// TIA Portal V17 export
// export: Created 2025-07-10T12:23:13.1481267Z, ExportSetting WithDefaults, DisplayName Totally Integrated Automation Portal, DisplayVersion V17, DisplayName TIA Portal Openness, DisplayVersion V17, DisplayName TIA Portal Version Control Interface, DisplayVersion V17, DisplayName SINAMICS Startdrive Advanced, DisplayVersion V17, DisplayName SINAMICS Startdrive G130, G150, S120, S150, SINAMICS MV, S210, DisplayVersion V17, DisplayName SINAMICS Startdrive G110M, G120, G120C, G120D, G120P, G115D, DisplayVersion V17, DisplayName STEP 7 Professional, DisplayVersion V17, DisplayName STEP 7 Safety, DisplayVersion V17, DisplayName WinCC Professional, DisplayVersion V17
FUNCTION_BLOCK "PR_PC4005_Operator_DecisionV4_77a371"   // FB1, LAD
VERSION : 0.1
// stored: AutoNumber true, IsIECCheckEnabled false, UDAEnableTagReadback false
   VAR_INPUT
      iAutoRunning : Bool;
      iOperatorAuthorizationPB : Bool;
      iPCAckZero : Bool;
      iPCBypass : Bool;
      iPCDataReadOver : Bool;
      iPCDataWriteOver : Bool;
      iPalletPresentAtStation : Bool;
      iProcessOver : Bool;
      iProcessStartFormPZR : Bool;
      iRejectPB : Bool;
      iResetMem : Bool;
      iReset_fault : Bool;
      iScanOver : Bool;
      iScanResultNok : Bool;
      iScanResultOk : Bool;
      iScannerBypass : Bool;
      iSstMode : Bool;
      iSstPB : Bool;
      iUnloadCycleSelection : Bool;
   END_VAR
   VAR_OUTPUT
      qPCReadCmd : Bool;
      qPCWriteCmd : Bool;
      qProcessOver : Bool;
      qResetPalletStatusData : Bool;
      qScanCmd : Bool;
   END_VAR
   VAR DB_SPECIFIC
      StateNo : Int;
      s29_WaitProcStart : Bool;
      s29_WaitProcStart_T1 : Bool;
      s30_WaitCartnSheetOp : Bool;
      s30_WaitCartnSheetOp_T1 : Bool;
      s31_ChkCycleSelect : Bool;
      s31_ChkCycleSelect_T1 : Bool;
      s31_ChkCycleSelect_T2 : Bool;
      s32_WaitScanOver : Bool;
      s32_WaitScanOver_T1 : Bool;
      s33_ChkScanResult : Bool;
      s33_ChkScanResult_T1 : Bool;
      s33_ChkScanResult_T2 : Bool;
      s34_WaitOpDecision : Bool;
      s34_WaitOpDecision_T1 : Bool;
      s34_WaitOpDecision_T2 : Bool;
      s35_ChkPCAckReset0 : Bool;
      s35_ChkPCAckReset0_T1 : Bool;
      s36_WaitDataReadPC : Bool;
      s36_WaitDataReadPC_T1 : Bool;
      s38_WaitProcStartLow : Bool;
      s38_WaitProcStartLow_T1 : Bool;
      s39_WaitPalletAbsnt : Bool;
      s39_WaitPalletAbsnt_T1 : Bool;
      s40_WaitFaultReset : Bool;
      s40_WaitFaultReset_T1 : Bool;
      s41_ChkPCAckReset0Up : Bool;
      s41_ChkPCAckReset0Up_T1 : Bool;
      s42_WaitDataUploadPC : Bool;
      s42_WaitDataUploadPC_T1 : Bool;
      s43_ChkRecovery : Bool;
      s43_ChkRecovery_T1 : Bool;
      s43_ChkRecovery_T2 : Bool;
      sPalletAccepted : Bool;
      sProcessOver : Bool;
      sSst : Bool;
      sSstPulse : Bool;
      sSstRise : Bool;
      sStWtResetRel : Bool;
      sStWtResetRel_T1 : Bool;
   END_VAR
   VAR_TEMP
      tOne : Bool;
   END_VAR
   VAR_TEMP   // added for the SCL form of the ladder/FBD networks
      _w1 : Bool;
   END_VAR
BEGIN

REGION Network 1
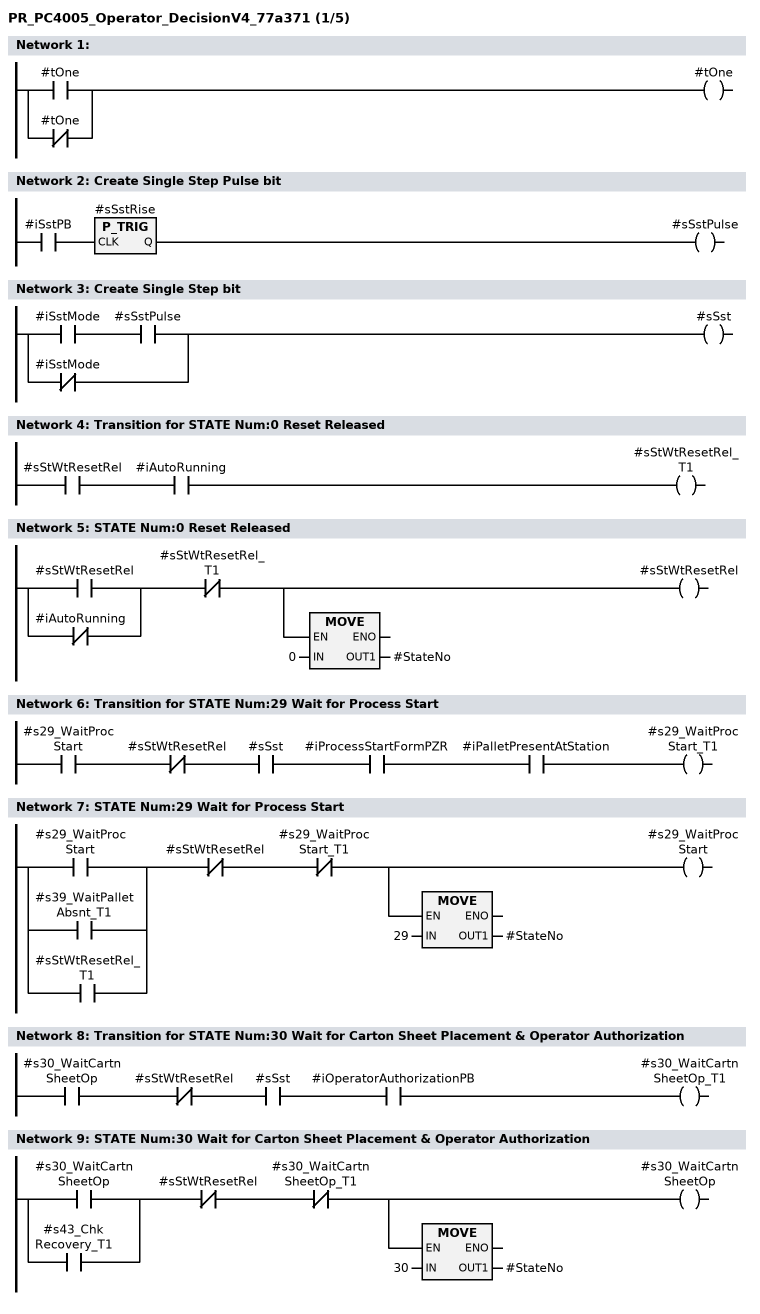
   RUNG wire#powerrail
      Contact( #tOne )
      wire#w1
      Coil( #tOne )
   END_RUNG
   RUNG wire#powerrail
      I_Contact( #tOne )
   END_RUNG wire#w1
   // the same network as SCL:
   #tOne := #tOne OR NOT #tOne;
END_REGION

REGION Network 2: Create Single Step Pulse bit
   RUNG wire#powerrail
      Contact( #iSstPB )
      P_Trig( #sSstRise )
      Coil( #sSstPulse )
   END_RUNG
   // the same network as SCL:
   #_w1 := #iSstPB AND NOT #sSstRise;   // rising edge
   #sSstRise := #iSstPB;
   #sSstPulse := #_w1;
END_REGION

REGION Network 3: Create Single Step bit
   RUNG wire#powerrail
      Contact( #iSstMode )
      Contact( #sSstPulse )
      wire#w1
      Coil( #sSst )
   END_RUNG
   RUNG wire#powerrail
      I_Contact( #iSstMode )
   END_RUNG wire#w1
   // the same network as SCL:
   #sSst := (#iSstMode AND #sSstPulse) OR NOT #iSstMode;
END_REGION

REGION Network 4: Transition for STATE Num:0 Reset Released
   RUNG wire#powerrail
      Contact( #sStWtResetRel )
      Contact( #iAutoRunning )
      Coil( #sStWtResetRel_T1 )
   END_RUNG
   // the same network as SCL:
   #sStWtResetRel_T1 := #sStWtResetRel AND #iAutoRunning;
END_REGION

REGION Network 5: STATE Num:0 Reset Released
   RUNG wire#powerrail
      Contact( #sStWtResetRel )
      wire#w1
      I_Contact( #sStWtResetRel_T1 )
      wire#w2
      Coil( #sStWtResetRel )
   END_RUNG
   RUNG wire#powerrail
      I_Contact( #iAutoRunning )
   END_RUNG wire#w1
   RUNG wire#w2
      { S7_GenerateENO := "TRUE" } Move(in := 0, out1 => #StateNo)
   END_RUNG
   // the same network as SCL:
   #sStWtResetRel := (#sStWtResetRel OR NOT #iAutoRunning) AND NOT #sStWtResetRel_T1;
   IF #sStWtResetRel THEN #StateNo := 0; END_IF;
END_REGION

REGION Network 6: Transition for STATE Num:29 Wait for Process Start
   RUNG wire#powerrail
      Contact( #s29_WaitProcStart )
      I_Contact( #sStWtResetRel )
      Contact( #sSst )
      Contact( #iProcessStartFormPZR )
      Contact( #iPalletPresentAtStation )
      Coil( #s29_WaitProcStart_T1 )
   END_RUNG
   // the same network as SCL:
   #s29_WaitProcStart_T1 := #s29_WaitProcStart AND NOT #sStWtResetRel AND #sSst AND #iProcessStartFormPZR AND #iPalletPresentAtStation;
END_REGION

REGION Network 7: STATE Num:29 Wait for Process Start
   RUNG wire#powerrail
      Contact( #s29_WaitProcStart )
      wire#w1
      I_Contact( #sStWtResetRel )
      I_Contact( #s29_WaitProcStart_T1 )
      wire#w2
      Coil( #s29_WaitProcStart )
   END_RUNG
   RUNG wire#powerrail
      Contact( #s39_WaitPalletAbsnt_T1 )
   END_RUNG wire#w1
   RUNG wire#powerrail
      Contact( #sStWtResetRel_T1 )
   END_RUNG wire#w1
   RUNG wire#w2
      { S7_GenerateENO := "TRUE" } Move(in := 29, out1 => #StateNo)
   END_RUNG
   // the same network as SCL:
   #s29_WaitProcStart := (#s29_WaitProcStart OR #s39_WaitPalletAbsnt_T1 OR #sStWtResetRel_T1) AND NOT #sStWtResetRel AND NOT #s29_WaitProcStart_T1;
   IF #s29_WaitProcStart THEN #StateNo := 29; END_IF;
END_REGION

REGION Network 8: Transition for STATE Num:30 Wait for Carton Sheet Placement & Operator Authorization
   RUNG wire#powerrail
      Contact( #s30_WaitCartnSheetOp )
      I_Contact( #sStWtResetRel )
      Contact( #sSst )
      Contact( #iOperatorAuthorizationPB )
      Coil( #s30_WaitCartnSheetOp_T1 )
   END_RUNG
   // the same network as SCL:
   #s30_WaitCartnSheetOp_T1 := #s30_WaitCartnSheetOp AND NOT #sStWtResetRel AND #sSst AND #iOperatorAuthorizationPB;
END_REGION

REGION Network 9: STATE Num:30 Wait for Carton Sheet Placement & Operator Authorization
   RUNG wire#powerrail
      Contact( #s30_WaitCartnSheetOp )
      wire#w1
      I_Contact( #sStWtResetRel )
      I_Contact( #s30_WaitCartnSheetOp_T1 )
      wire#w2
      Coil( #s30_WaitCartnSheetOp )
   END_RUNG
   RUNG wire#powerrail
      Contact( #s43_ChkRecovery_T1 )
   END_RUNG wire#w1
   RUNG wire#w2
      { S7_GenerateENO := "TRUE" } Move(in := 30, out1 => #StateNo)
   END_RUNG
   // the same network as SCL:
   #s30_WaitCartnSheetOp := (#s30_WaitCartnSheetOp OR #s43_ChkRecovery_T1) AND NOT #sStWtResetRel AND NOT #s30_WaitCartnSheetOp_T1;
   IF #s30_WaitCartnSheetOp THEN #StateNo := 30; END_IF;
END_REGION

REGION Network 10: Transition for STATE Num:31 Check Cycle Selection
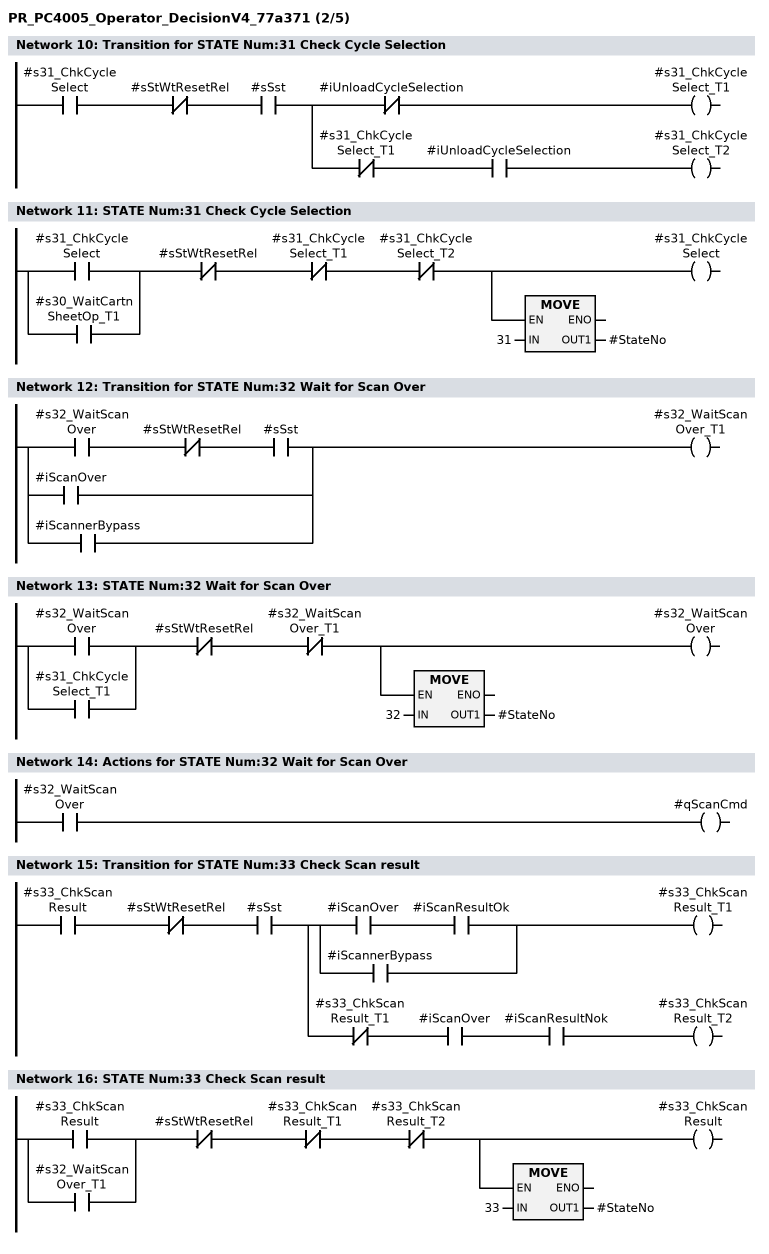
   RUNG wire#powerrail
      Contact( #s31_ChkCycleSelect )
      I_Contact( #sStWtResetRel )
      Contact( #sSst )
      wire#w1
      I_Contact( #iUnloadCycleSelection )
      Coil( #s31_ChkCycleSelect_T1 )
   END_RUNG
   RUNG wire#w1
      I_Contact( #s31_ChkCycleSelect_T1 )
      Contact( #iUnloadCycleSelection )
      Coil( #s31_ChkCycleSelect_T2 )
   END_RUNG
   // the same network as SCL:
   #_w1 := #s31_ChkCycleSelect AND NOT #sStWtResetRel AND #sSst;
   #s31_ChkCycleSelect_T1 := #_w1 AND NOT #iUnloadCycleSelection;
   #s31_ChkCycleSelect_T2 := #_w1 AND NOT #s31_ChkCycleSelect_T1 AND #iUnloadCycleSelection;
END_REGION

REGION Network 11: STATE Num:31 Check Cycle Selection
   RUNG wire#powerrail
      Contact( #s31_ChkCycleSelect )
      wire#w1
      I_Contact( #sStWtResetRel )
      I_Contact( #s31_ChkCycleSelect_T1 )
      I_Contact( #s31_ChkCycleSelect_T2 )
      wire#w2
      Coil( #s31_ChkCycleSelect )
   END_RUNG
   RUNG wire#powerrail
      Contact( #s30_WaitCartnSheetOp_T1 )
   END_RUNG wire#w1
   RUNG wire#w2
      { S7_GenerateENO := "TRUE" } Move(in := 31, out1 => #StateNo)
   END_RUNG
   // the same network as SCL:
   #s31_ChkCycleSelect := (#s31_ChkCycleSelect OR #s30_WaitCartnSheetOp_T1) AND NOT #sStWtResetRel AND NOT #s31_ChkCycleSelect_T1 AND NOT #s31_ChkCycleSelect_T2;
   IF #s31_ChkCycleSelect THEN #StateNo := 31; END_IF;
END_REGION

REGION Network 12: Transition for STATE Num:32 Wait for Scan Over
   RUNG wire#powerrail
      Contact( #s32_WaitScanOver )
      I_Contact( #sStWtResetRel )
      Contact( #sSst )
      wire#w1
      Coil( #s32_WaitScanOver_T1 )
   END_RUNG
   RUNG wire#powerrail
      Contact( #iScanOver )
   END_RUNG wire#w1
   RUNG wire#powerrail
      Contact( #iScannerBypass )
   END_RUNG wire#w1
   // the same network as SCL:
   #s32_WaitScanOver_T1 := (#s32_WaitScanOver AND NOT #sStWtResetRel AND #sSst) OR #iScanOver OR #iScannerBypass;
END_REGION

REGION Network 13: STATE Num:32 Wait for Scan Over
   RUNG wire#powerrail
      Contact( #s32_WaitScanOver )
      wire#w1
      I_Contact( #sStWtResetRel )
      I_Contact( #s32_WaitScanOver_T1 )
      wire#w2
      Coil( #s32_WaitScanOver )
   END_RUNG
   RUNG wire#powerrail
      Contact( #s31_ChkCycleSelect_T1 )
   END_RUNG wire#w1
   RUNG wire#w2
      { S7_GenerateENO := "TRUE" } Move(in := 32, out1 => #StateNo)
   END_RUNG
   // the same network as SCL:
   #s32_WaitScanOver := (#s32_WaitScanOver OR #s31_ChkCycleSelect_T1) AND NOT #sStWtResetRel AND NOT #s32_WaitScanOver_T1;
   IF #s32_WaitScanOver THEN #StateNo := 32; END_IF;
END_REGION

REGION Network 14: Actions for STATE Num:32 Wait for Scan Over
   RUNG wire#powerrail
      Contact( #s32_WaitScanOver )
      Coil( #qScanCmd )
   END_RUNG
   // the same network as SCL:
   #qScanCmd := #s32_WaitScanOver;
END_REGION

REGION Network 15: Transition for STATE Num:33 Check Scan result
   RUNG wire#powerrail
      Contact( #s33_ChkScanResult )
      I_Contact( #sStWtResetRel )
      Contact( #sSst )
      wire#w1
      Contact( #iScanOver )
      Contact( #iScanResultOk )
      wire#w2
      Coil( #s33_ChkScanResult_T1 )
   END_RUNG
   RUNG wire#w1
      Contact( #iScannerBypass )
   END_RUNG wire#w2
   RUNG wire#w1
      I_Contact( #s33_ChkScanResult_T1 )
      Contact( #iScanOver )
      Contact( #iScanResultNok )
      Coil( #s33_ChkScanResult_T2 )
   END_RUNG
   // the same network as SCL:
   #_w1 := #s33_ChkScanResult AND NOT #sStWtResetRel AND #sSst;
   #s33_ChkScanResult_T1 := #_w1 AND ((#iScanOver AND #iScanResultOk) OR #iScannerBypass);
   #s33_ChkScanResult_T2 := #_w1 AND NOT #s33_ChkScanResult_T1 AND #iScanOver AND #iScanResultNok;
END_REGION

REGION Network 16: STATE Num:33 Check Scan result
   RUNG wire#powerrail
      Contact( #s33_ChkScanResult )
      wire#w1
      I_Contact( #sStWtResetRel )
      I_Contact( #s33_ChkScanResult_T1 )
      I_Contact( #s33_ChkScanResult_T2 )
      wire#w2
      Coil( #s33_ChkScanResult )
   END_RUNG
   RUNG wire#powerrail
      Contact( #s32_WaitScanOver_T1 )
   END_RUNG wire#w1
   RUNG wire#w2
      { S7_GenerateENO := "TRUE" } Move(in := 33, out1 => #StateNo)
   END_RUNG
   // the same network as SCL:
   #s33_ChkScanResult := (#s33_ChkScanResult OR #s32_WaitScanOver_T1) AND NOT #sStWtResetRel AND NOT #s33_ChkScanResult_T1 AND NOT #s33_ChkScanResult_T2;
   IF #s33_ChkScanResult THEN #StateNo := 33; END_IF;
END_REGION

REGION Network 17: Transition for STATE Num:34 Wait for Operator Decision
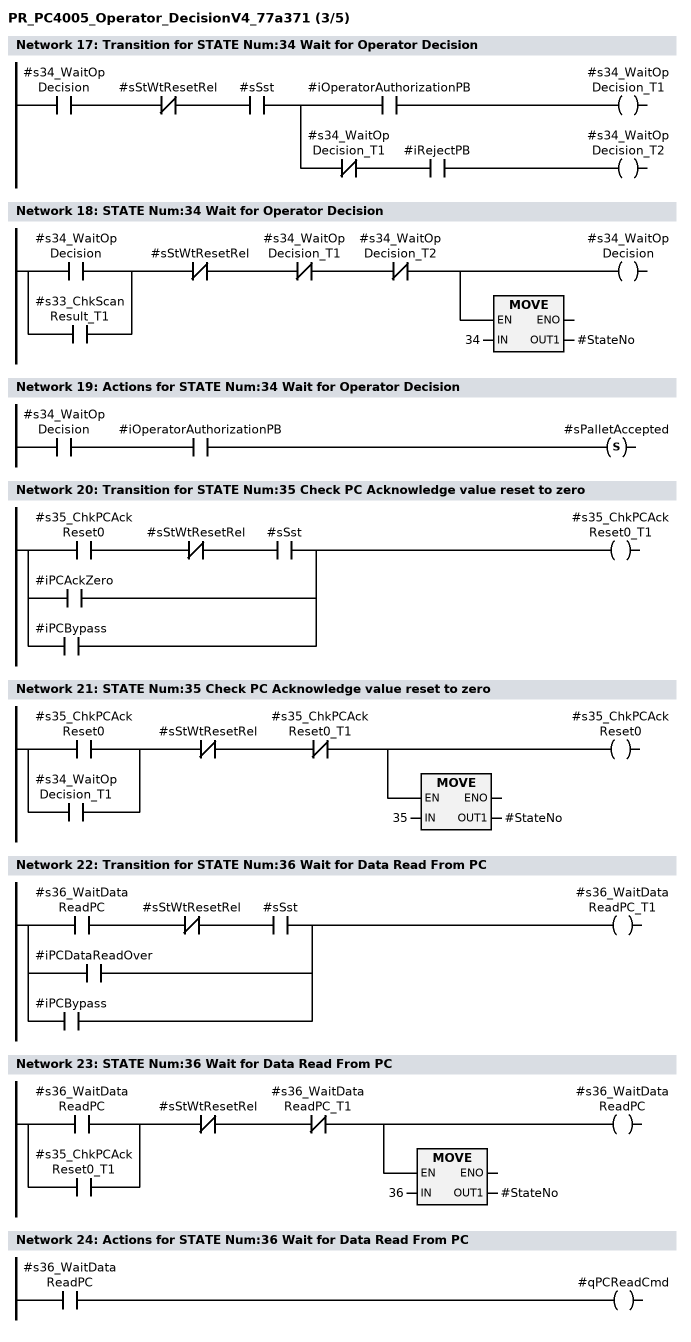
   RUNG wire#powerrail
      Contact( #s34_WaitOpDecision )
      I_Contact( #sStWtResetRel )
      Contact( #sSst )
      wire#w1
      Contact( #iOperatorAuthorizationPB )
      Coil( #s34_WaitOpDecision_T1 )
   END_RUNG
   RUNG wire#w1
      I_Contact( #s34_WaitOpDecision_T1 )
      Contact( #iRejectPB )
      Coil( #s34_WaitOpDecision_T2 )
   END_RUNG
   // the same network as SCL:
   #_w1 := #s34_WaitOpDecision AND NOT #sStWtResetRel AND #sSst;
   #s34_WaitOpDecision_T1 := #_w1 AND #iOperatorAuthorizationPB;
   #s34_WaitOpDecision_T2 := #_w1 AND NOT #s34_WaitOpDecision_T1 AND #iRejectPB;
END_REGION

REGION Network 18: STATE Num:34 Wait for Operator Decision
   RUNG wire#powerrail
      Contact( #s34_WaitOpDecision )
      wire#w1
      I_Contact( #sStWtResetRel )
      I_Contact( #s34_WaitOpDecision_T1 )
      I_Contact( #s34_WaitOpDecision_T2 )
      wire#w2
      Coil( #s34_WaitOpDecision )
   END_RUNG
   RUNG wire#powerrail
      Contact( #s33_ChkScanResult_T1 )
   END_RUNG wire#w1
   RUNG wire#w2
      { S7_GenerateENO := "TRUE" } Move(in := 34, out1 => #StateNo)
   END_RUNG
   // the same network as SCL:
   #s34_WaitOpDecision := (#s34_WaitOpDecision OR #s33_ChkScanResult_T1) AND NOT #sStWtResetRel AND NOT #s34_WaitOpDecision_T1 AND NOT #s34_WaitOpDecision_T2;
   IF #s34_WaitOpDecision THEN #StateNo := 34; END_IF;
END_REGION

REGION Network 19: Actions for STATE Num:34 Wait for Operator Decision
   RUNG wire#powerrail
      Contact( #s34_WaitOpDecision )
      Contact( #iOperatorAuthorizationPB )
      S_Coil( #sPalletAccepted )
   END_RUNG
   // the same network as SCL:
   IF #s34_WaitOpDecision AND #iOperatorAuthorizationPB THEN #sPalletAccepted := TRUE; END_IF;
END_REGION

REGION Network 20: Transition for STATE Num:35 Check PC Acknowledge value reset to zero
   RUNG wire#powerrail
      Contact( #s35_ChkPCAckReset0 )
      I_Contact( #sStWtResetRel )
      Contact( #sSst )
      wire#w1
      Coil( #s35_ChkPCAckReset0_T1 )
   END_RUNG
   RUNG wire#powerrail
      Contact( #iPCAckZero )
   END_RUNG wire#w1
   RUNG wire#powerrail
      Contact( #iPCBypass )
   END_RUNG wire#w1
   // the same network as SCL:
   #s35_ChkPCAckReset0_T1 := (#s35_ChkPCAckReset0 AND NOT #sStWtResetRel AND #sSst) OR #iPCAckZero OR #iPCBypass;
END_REGION

REGION Network 21: STATE Num:35 Check PC Acknowledge value reset to zero
   RUNG wire#powerrail
      Contact( #s35_ChkPCAckReset0 )
      wire#w1
      I_Contact( #sStWtResetRel )
      I_Contact( #s35_ChkPCAckReset0_T1 )
      wire#w2
      Coil( #s35_ChkPCAckReset0 )
   END_RUNG
   RUNG wire#powerrail
      Contact( #s34_WaitOpDecision_T1 )
   END_RUNG wire#w1
   RUNG wire#w2
      { S7_GenerateENO := "TRUE" } Move(in := 35, out1 => #StateNo)
   END_RUNG
   // the same network as SCL:
   #s35_ChkPCAckReset0 := (#s35_ChkPCAckReset0 OR #s34_WaitOpDecision_T1) AND NOT #sStWtResetRel AND NOT #s35_ChkPCAckReset0_T1;
   IF #s35_ChkPCAckReset0 THEN #StateNo := 35; END_IF;
END_REGION

REGION Network 22: Transition for STATE Num:36 Wait for Data Read From PC
   RUNG wire#powerrail
      Contact( #s36_WaitDataReadPC )
      I_Contact( #sStWtResetRel )
      Contact( #sSst )
      wire#w1
      Coil( #s36_WaitDataReadPC_T1 )
   END_RUNG
   RUNG wire#powerrail
      Contact( #iPCDataReadOver )
   END_RUNG wire#w1
   RUNG wire#powerrail
      Contact( #iPCBypass )
   END_RUNG wire#w1
   // the same network as SCL:
   #s36_WaitDataReadPC_T1 := (#s36_WaitDataReadPC AND NOT #sStWtResetRel AND #sSst) OR #iPCDataReadOver OR #iPCBypass;
END_REGION

REGION Network 23: STATE Num:36 Wait for Data Read From PC
   RUNG wire#powerrail
      Contact( #s36_WaitDataReadPC )
      wire#w1
      I_Contact( #sStWtResetRel )
      I_Contact( #s36_WaitDataReadPC_T1 )
      wire#w2
      Coil( #s36_WaitDataReadPC )
   END_RUNG
   RUNG wire#powerrail
      Contact( #s35_ChkPCAckReset0_T1 )
   END_RUNG wire#w1
   RUNG wire#w2
      { S7_GenerateENO := "TRUE" } Move(in := 36, out1 => #StateNo)
   END_RUNG
   // the same network as SCL:
   #s36_WaitDataReadPC := (#s36_WaitDataReadPC OR #s35_ChkPCAckReset0_T1) AND NOT #sStWtResetRel AND NOT #s36_WaitDataReadPC_T1;
   IF #s36_WaitDataReadPC THEN #StateNo := 36; END_IF;
END_REGION

REGION Network 24: Actions for STATE Num:36 Wait for Data Read From PC
   RUNG wire#powerrail
      Contact( #s36_WaitDataReadPC )
      Coil( #qPCReadCmd )
   END_RUNG
   // the same network as SCL:
   #qPCReadCmd := #s36_WaitDataReadPC;
END_REGION

REGION Network 25: Transition for STATE Num:38 Wait for Process Start Low
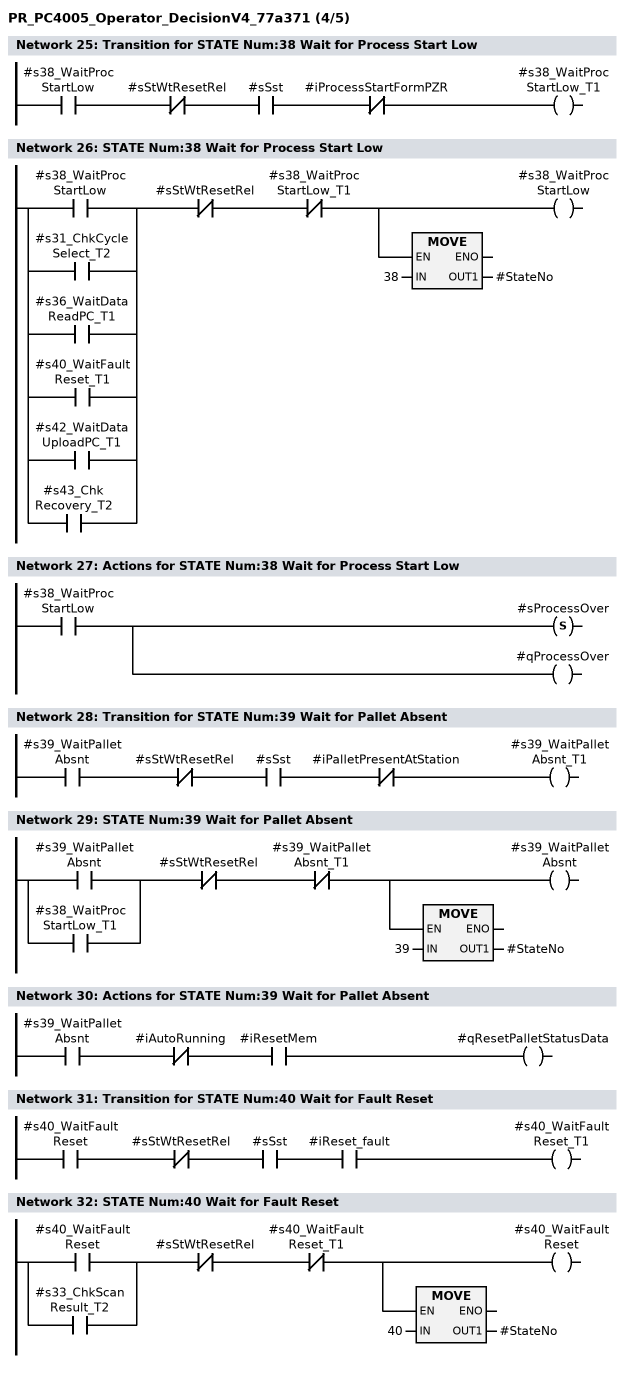
   RUNG wire#powerrail
      Contact( #s38_WaitProcStartLow )
      I_Contact( #sStWtResetRel )
      Contact( #sSst )
      I_Contact( #iProcessStartFormPZR )
      Coil( #s38_WaitProcStartLow_T1 )
   END_RUNG
   // the same network as SCL:
   #s38_WaitProcStartLow_T1 := #s38_WaitProcStartLow AND NOT #sStWtResetRel AND #sSst AND NOT #iProcessStartFormPZR;
END_REGION

REGION Network 26: STATE Num:38 Wait for Process Start Low
   RUNG wire#powerrail
      Contact( #s38_WaitProcStartLow )
      wire#w1
      I_Contact( #sStWtResetRel )
      I_Contact( #s38_WaitProcStartLow_T1 )
      wire#w2
      Coil( #s38_WaitProcStartLow )
   END_RUNG
   RUNG wire#powerrail
      Contact( #s31_ChkCycleSelect_T2 )
   END_RUNG wire#w1
   RUNG wire#powerrail
      Contact( #s36_WaitDataReadPC_T1 )
   END_RUNG wire#w1
   RUNG wire#powerrail
      Contact( #s40_WaitFaultReset_T1 )
   END_RUNG wire#w1
   RUNG wire#powerrail
      Contact( #s42_WaitDataUploadPC_T1 )
   END_RUNG wire#w1
   RUNG wire#powerrail
      Contact( #s43_ChkRecovery_T2 )
   END_RUNG wire#w1
   RUNG wire#w2
      { S7_GenerateENO := "TRUE" } Move(in := 38, out1 => #StateNo)
   END_RUNG
   // the same network as SCL:
   #s38_WaitProcStartLow := (#s38_WaitProcStartLow OR #s31_ChkCycleSelect_T2 OR #s36_WaitDataReadPC_T1 OR #s40_WaitFaultReset_T1 OR #s42_WaitDataUploadPC_T1 OR #s43_ChkRecovery_T2) AND NOT #sStWtResetRel AND NOT #s38_WaitProcStartLow_T1;
   IF #s38_WaitProcStartLow THEN #StateNo := 38; END_IF;
END_REGION

REGION Network 27: Actions for STATE Num:38 Wait for Process Start Low
   RUNG wire#powerrail
      Contact( #s38_WaitProcStartLow )
      wire#w1
      S_Coil( #sProcessOver )
   END_RUNG
   RUNG wire#w1
      Coil( #qProcessOver )
   END_RUNG
   // the same network as SCL:
   IF #s38_WaitProcStartLow THEN #sProcessOver := TRUE; END_IF;
   #qProcessOver := #s38_WaitProcStartLow;
END_REGION

REGION Network 28: Transition for STATE Num:39 Wait for Pallet Absent
   RUNG wire#powerrail
      Contact( #s39_WaitPalletAbsnt )
      I_Contact( #sStWtResetRel )
      Contact( #sSst )
      I_Contact( #iPalletPresentAtStation )
      Coil( #s39_WaitPalletAbsnt_T1 )
   END_RUNG
   // the same network as SCL:
   #s39_WaitPalletAbsnt_T1 := #s39_WaitPalletAbsnt AND NOT #sStWtResetRel AND #sSst AND NOT #iPalletPresentAtStation;
END_REGION

REGION Network 29: STATE Num:39 Wait for Pallet Absent
   RUNG wire#powerrail
      Contact( #s39_WaitPalletAbsnt )
      wire#w1
      I_Contact( #sStWtResetRel )
      I_Contact( #s39_WaitPalletAbsnt_T1 )
      wire#w2
      Coil( #s39_WaitPalletAbsnt )
   END_RUNG
   RUNG wire#powerrail
      Contact( #s38_WaitProcStartLow_T1 )
   END_RUNG wire#w1
   RUNG wire#w2
      { S7_GenerateENO := "TRUE" } Move(in := 39, out1 => #StateNo)
   END_RUNG
   // the same network as SCL:
   #s39_WaitPalletAbsnt := (#s39_WaitPalletAbsnt OR #s38_WaitProcStartLow_T1) AND NOT #sStWtResetRel AND NOT #s39_WaitPalletAbsnt_T1;
   IF #s39_WaitPalletAbsnt THEN #StateNo := 39; END_IF;
END_REGION

REGION Network 30: Actions for STATE Num:39 Wait for Pallet Absent
   RUNG wire#powerrail
      Contact( #s39_WaitPalletAbsnt )
      I_Contact( #iAutoRunning )
      Contact( #iResetMem )
      Coil( #qResetPalletStatusData )
   END_RUNG
   // the same network as SCL:
   #qResetPalletStatusData := #s39_WaitPalletAbsnt AND NOT #iAutoRunning AND #iResetMem;
END_REGION

REGION Network 31: Transition for STATE Num:40 Wait for Fault Reset
   RUNG wire#powerrail
      Contact( #s40_WaitFaultReset )
      I_Contact( #sStWtResetRel )
      Contact( #sSst )
      Contact( #iReset_fault )
      Coil( #s40_WaitFaultReset_T1 )
   END_RUNG
   // the same network as SCL:
   #s40_WaitFaultReset_T1 := #s40_WaitFaultReset AND NOT #sStWtResetRel AND #sSst AND #iReset_fault;
END_REGION

REGION Network 32: STATE Num:40 Wait for Fault Reset
   RUNG wire#powerrail
      Contact( #s40_WaitFaultReset )
      wire#w1
      I_Contact( #sStWtResetRel )
      I_Contact( #s40_WaitFaultReset_T1 )
      wire#w2
      Coil( #s40_WaitFaultReset )
   END_RUNG
   RUNG wire#powerrail
      Contact( #s33_ChkScanResult_T2 )
   END_RUNG wire#w1
   RUNG wire#w2
      { S7_GenerateENO := "TRUE" } Move(in := 40, out1 => #StateNo)
   END_RUNG
   // the same network as SCL:
   #s40_WaitFaultReset := (#s40_WaitFaultReset OR #s33_ChkScanResult_T2) AND NOT #sStWtResetRel AND NOT #s40_WaitFaultReset_T1;
   IF #s40_WaitFaultReset THEN #StateNo := 40; END_IF;
END_REGION

REGION Network 33: Transition for STATE Num:41 Check PC Acknowledge value reset to zero for Upload
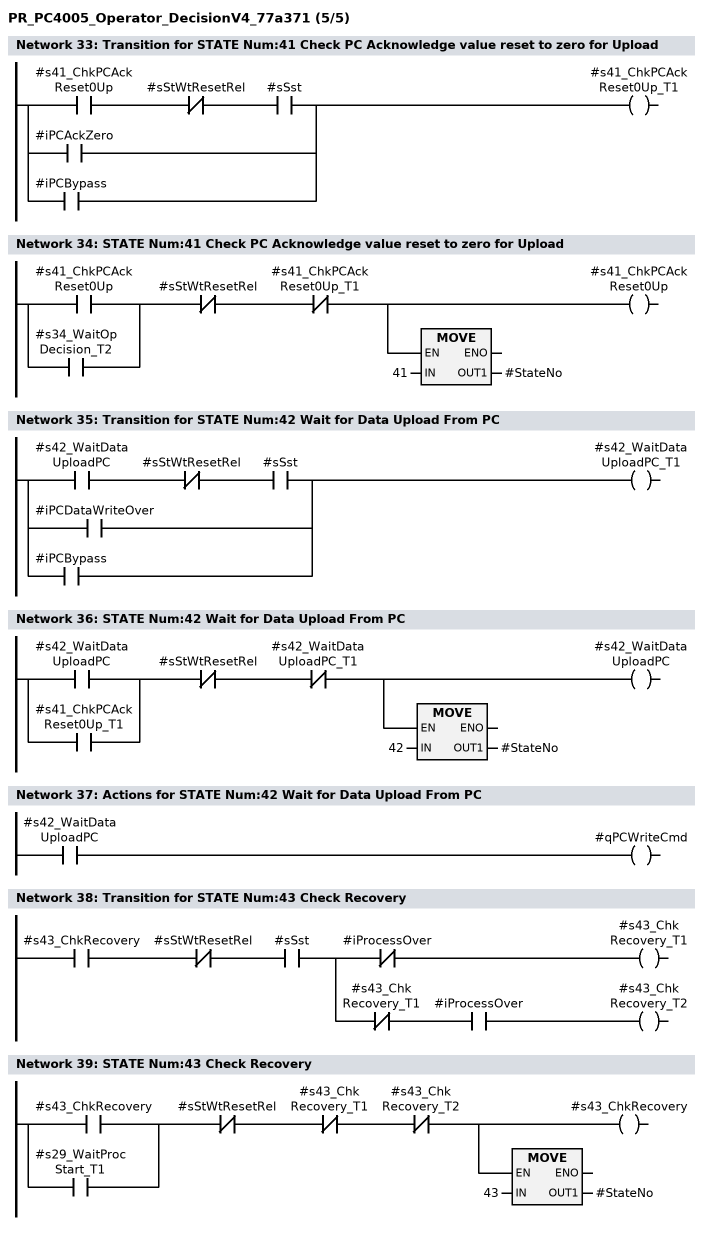
   RUNG wire#powerrail
      Contact( #s41_ChkPCAckReset0Up )
      I_Contact( #sStWtResetRel )
      Contact( #sSst )
      wire#w1
      Coil( #s41_ChkPCAckReset0Up_T1 )
   END_RUNG
   RUNG wire#powerrail
      Contact( #iPCAckZero )
   END_RUNG wire#w1
   RUNG wire#powerrail
      Contact( #iPCBypass )
   END_RUNG wire#w1
   // the same network as SCL:
   #s41_ChkPCAckReset0Up_T1 := (#s41_ChkPCAckReset0Up AND NOT #sStWtResetRel AND #sSst) OR #iPCAckZero OR #iPCBypass;
END_REGION

REGION Network 34: STATE Num:41 Check PC Acknowledge value reset to zero for Upload
   RUNG wire#powerrail
      Contact( #s41_ChkPCAckReset0Up )
      wire#w1
      I_Contact( #sStWtResetRel )
      I_Contact( #s41_ChkPCAckReset0Up_T1 )
      wire#w2
      Coil( #s41_ChkPCAckReset0Up )
   END_RUNG
   RUNG wire#powerrail
      Contact( #s34_WaitOpDecision_T2 )
   END_RUNG wire#w1
   RUNG wire#w2
      { S7_GenerateENO := "TRUE" } Move(in := 41, out1 => #StateNo)
   END_RUNG
   // the same network as SCL:
   #s41_ChkPCAckReset0Up := (#s41_ChkPCAckReset0Up OR #s34_WaitOpDecision_T2) AND NOT #sStWtResetRel AND NOT #s41_ChkPCAckReset0Up_T1;
   IF #s41_ChkPCAckReset0Up THEN #StateNo := 41; END_IF;
END_REGION

REGION Network 35: Transition for STATE Num:42 Wait for Data Upload From PC
   RUNG wire#powerrail
      Contact( #s42_WaitDataUploadPC )
      I_Contact( #sStWtResetRel )
      Contact( #sSst )
      wire#w1
      Coil( #s42_WaitDataUploadPC_T1 )
   END_RUNG
   RUNG wire#powerrail
      Contact( #iPCDataWriteOver )
   END_RUNG wire#w1
   RUNG wire#powerrail
      Contact( #iPCBypass )
   END_RUNG wire#w1
   // the same network as SCL:
   #s42_WaitDataUploadPC_T1 := (#s42_WaitDataUploadPC AND NOT #sStWtResetRel AND #sSst) OR #iPCDataWriteOver OR #iPCBypass;
END_REGION

REGION Network 36: STATE Num:42 Wait for Data Upload From PC
   RUNG wire#powerrail
      Contact( #s42_WaitDataUploadPC )
      wire#w1
      I_Contact( #sStWtResetRel )
      I_Contact( #s42_WaitDataUploadPC_T1 )
      wire#w2
      Coil( #s42_WaitDataUploadPC )
   END_RUNG
   RUNG wire#powerrail
      Contact( #s41_ChkPCAckReset0Up_T1 )
   END_RUNG wire#w1
   RUNG wire#w2
      { S7_GenerateENO := "TRUE" } Move(in := 42, out1 => #StateNo)
   END_RUNG
   // the same network as SCL:
   #s42_WaitDataUploadPC := (#s42_WaitDataUploadPC OR #s41_ChkPCAckReset0Up_T1) AND NOT #sStWtResetRel AND NOT #s42_WaitDataUploadPC_T1;
   IF #s42_WaitDataUploadPC THEN #StateNo := 42; END_IF;
END_REGION

REGION Network 37: Actions for STATE Num:42 Wait for Data Upload From PC
   RUNG wire#powerrail
      Contact( #s42_WaitDataUploadPC )
      Coil( #qPCWriteCmd )
   END_RUNG
   // the same network as SCL:
   #qPCWriteCmd := #s42_WaitDataUploadPC;
END_REGION

REGION Network 38: Transition for STATE Num:43 Check Recovery
   RUNG wire#powerrail
      Contact( #s43_ChkRecovery )
      I_Contact( #sStWtResetRel )
      Contact( #sSst )
      wire#w1
      I_Contact( #iProcessOver )
      Coil( #s43_ChkRecovery_T1 )
   END_RUNG
   RUNG wire#w1
      I_Contact( #s43_ChkRecovery_T1 )
      Contact( #iProcessOver )
      Coil( #s43_ChkRecovery_T2 )
   END_RUNG
   // the same network as SCL:
   #_w1 := #s43_ChkRecovery AND NOT #sStWtResetRel AND #sSst;
   #s43_ChkRecovery_T1 := #_w1 AND NOT #iProcessOver;
   #s43_ChkRecovery_T2 := #_w1 AND NOT #s43_ChkRecovery_T1 AND #iProcessOver;
END_REGION

REGION Network 39: STATE Num:43 Check Recovery
   RUNG wire#powerrail
      Contact( #s43_ChkRecovery )
      wire#w1
      I_Contact( #sStWtResetRel )
      I_Contact( #s43_ChkRecovery_T1 )
      I_Contact( #s43_ChkRecovery_T2 )
      wire#w2
      Coil( #s43_ChkRecovery )
   END_RUNG
   RUNG wire#powerrail
      Contact( #s29_WaitProcStart_T1 )
   END_RUNG wire#w1
   RUNG wire#w2
      { S7_GenerateENO := "TRUE" } Move(in := 43, out1 => #StateNo)
   END_RUNG
   // the same network as SCL:
   #s43_ChkRecovery := (#s43_ChkRecovery OR #s29_WaitProcStart_T1) AND NOT #sStWtResetRel AND NOT #s43_ChkRecovery_T1 AND NOT #s43_ChkRecovery_T2;
   IF #s43_ChkRecovery THEN #StateNo := 43; END_IF;
END_REGION
END_FUNCTION_BLOCK
